Fanuc KAREL source: kt00165.KL

-- PROVISIONAL review KL for V1013-1; original PC SHA256 130408e056c73dffc68a44d37e549ddb04700f3d838d1c05b4f81fe4777b3947
-- Incomplete behavior may be omitted. Consult companion uncertainty JSON. Do not deploy.
PROGRAM KT00165
%NOLOCKGROUP
VAR
  I1 : INTEGER
  OUT : INTEGER
-- UNRESOLVED_DECL Y2 type=002018
BEGIN
  -- UNRESOLVED_PC offsets 5-16; opcodes 2E,23
  -- UNRESOLVED_PC offsets 21-35; opcodes 2E,22,9D,33,B2
  -- UNRESOLVED_PC offsets 40-62; opcodes 21,22,9D,33,B1,56,23
  -- UNRESOLVED_PC offsets 67-71; opcodes 7F
END KT00165
